(* IEC 61131-3 sources: model-first-plc-agent-ai/results/T3-W-27, 2 files *)

(* ---- a1_code.st ---- *)
FUNCTION_BLOCK FB_TankRuntime
VAR_INPUT
    start : BOOL;
    stop : BOOL;
    LSH : BOOL;
    LSHH : BOOL;
    TON_Duration : TIME;
    TOF_Duration : TIME;
END_VAR
VAR_OUTPUT
    fill_valve : BOOL;
    discharge_valve : BOOL;
END_VAR
VAR
    state_id : INT := 0;
    previous_state : INT := 0;
    filling_active : BOOL := FALSE;
    ton_q : BOOL := FALSE;
    tof_q : BOOL := FALSE;
    fill_timer : TON;
    pause_timer : TOF;
END_VAR

(* Evaluate timers using the current filling-step activity. *)
filling_active := (state_id = 1);

fill_timer(IN := filling_active, PT := TON_Duration);
pause_timer(IN := filling_active, PT := TOF_Duration);

ton_q := fill_timer.Q;
tof_q := pause_timer.Q;

previous_state := state_id;

(* Evaluate transitions from the current situation. *)
CASE state_id OF
    0:
        IF start AND NOT stop AND NOT LSH AND NOT LSHH THEN
            state_id := 1;
        END_IF;

    1:
        IF stop OR LSH OR LSHH THEN
            state_id := 0;
        ELSIF ton_q AND NOT stop AND NOT LSH AND NOT LSHH THEN
            state_id := 2;
        END_IF;

    2:
        IF stop OR LSH OR LSHH THEN
            state_id := 0;
        ELSIF NOT tof_q AND NOT stop AND NOT LSH AND NOT LSHH THEN
            state_id := 1;
        END_IF;

ELSE
    state_id := 0;
END_CASE;

(* Synchronize timer inputs immediately with step entry or exit.
   In particular, the TOF falling edge occurs on entry to pause. *)
IF state_id <> previous_state THEN
    filling_active := (state_id = 1);

    fill_timer(IN := filling_active, PT := TON_Duration);
    pause_timer(IN := filling_active, PT := TOF_Duration);

    ton_q := fill_timer.Q;
    tof_q := pause_timer.Q;
END_IF;

(* Continuous actions of the resulting GRAFCET situation. *)
fill_valve := (state_id = 1);
discharge_valve := FALSE;

END_FUNCTION_BLOCK

PROGRAM Main
VAR
    StartCommand AT %IX100.0 : BOOL;
    StopCommand AT %IX100.1 : BOOL;
    LSH AT %IX100.2 : BOOL;
    LSHH AT %IX100.3 : BOOL;
    FillValve AT %QX100.0 : BOOL;
    DischargeValve AT %QX100.1 : BOOL;
END_VAR
VAR
    (* Adjustable timer parameters; defaults are commissioning values. *)
    TON_Duration : TIME := T#5s;
    TOF_Duration : TIME := T#5s;
    start_edge : R_TRIG;
    tank_runtime : FB_TankRuntime;
END_VAR

start_edge(CLK := StartCommand);

tank_runtime(
    start := start_edge.Q,
    stop := StopCommand,
    LSH := LSH,
    LSHH := LSHH,
    TON_Duration := TON_Duration,
    TOF_Duration := TOF_Duration
);

FillValve := tank_runtime.fill_valve;
DischargeValve := tank_runtime.discharge_valve;

END_PROGRAM

(* ---- a2_code.st ---- *)
FUNCTION_BLOCK FB_TankControl
VAR_INPUT
    StartCommand : BOOL;
    StopCommand : BOOL;
    LSH : BOOL;
    LSHH : BOOL;
    TON_Duration : TIME;
    TOF_Duration : TIME;
END_VAR
VAR_OUTPUT
    fill_valve : BOOL;
    discharge_valve : BOOL;
END_VAR
VAR
    sequence_state : INT := 0;
    start_edge : R_TRIG;
    filling_timer : TON;
    pause_timer : TOF;
    start : BOOL;
    stop : BOOL;
    ton_q : BOOL;
    tof_q : BOOL;
    filling_active : BOOL;
END_VAR

start_edge(CLK := StartCommand);
start := start_edge.Q;
stop := StopCommand;

filling_active := (sequence_state = 1);

filling_timer(
    IN := filling_active,
    PT := TON_Duration
);
pause_timer(
    IN := filling_active,
    PT := TOF_Duration
);

ton_q := filling_timer.Q;
tof_q := pause_timer.Q;

IF stop THEN
    sequence_state := 0;
ELSE
    CASE sequence_state OF
        0:
            IF start AND NOT LSH THEN
                sequence_state := 1;
            END_IF;

        1:
            IF LSH THEN
                sequence_state := 0;
            ELSIF ton_q THEN
                sequence_state := 2;
            END_IF;

        2:
            IF LSH THEN
                sequence_state := 0;
            ELSIF NOT tof_q THEN
                sequence_state := 1;
            END_IF;

        ELSE
            sequence_state := 0;
    END_CASE;
END_IF;

fill_valve := (sequence_state = 1) AND NOT stop;
discharge_valve := FALSE;

END_FUNCTION_BLOCK

PROGRAM Main
VAR
    StartCommand AT %IX100.0 : BOOL;
    StopCommand AT %IX100.1 : BOOL;
    LSH AT %IX100.2 : BOOL;
    LSHH AT %IX100.3 : BOOL;
    FillValve AT %QX100.0 : BOOL;
    DischargeValve AT %QX100.1 : BOOL;
END_VAR
VAR
    tank_controller : FB_TankControl;
    (* Configurable example presets; set to the required process values. *)
    TON_Duration : TIME := T#5s;
    TOF_Duration : TIME := T#5s;
END_VAR

tank_controller(
    StartCommand := StartCommand,
    StopCommand := StopCommand,
    LSH := LSH,
    LSHH := LSHH,
    TON_Duration := TON_Duration,
    TOF_Duration := TOF_Duration
);

FillValve := tank_controller.fill_valve;
DischargeValve := tank_controller.discharge_valve;

END_PROGRAM
